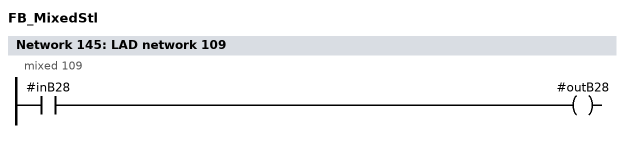
   RUNG wire#powerrail
      Contact( #inB28 )
      Coil( #outB28 )
   END_RUNG
   // the same network as SCL:
   #outB28 := #inB28;
END_REGION

REGION Network 146 (FBD): FBD network 110
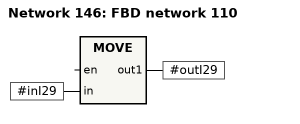
   #outI29 := #inI29;
END_REGION

REGION Network 147 (SCL): SCL network 111
   #tI10 := #inI30 + #cI20;
           IF #inB30 THEN
               #outR10 := #inR10 * 2.0;
           END_IF;
END_REGION

NETWORK
TITLE = STL network 37
      A     #inB36;
      AN    #stB36;
      =     #outB36;

REGION Network 149: LAD network 112
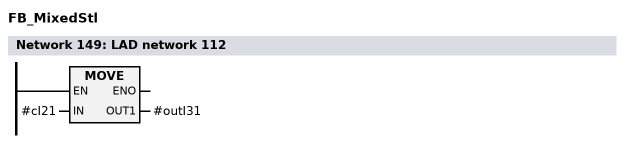
   RUNG wire#powerrail
      Move(in := #cI21, out1 => #outI31)
   END_RUNG
   // the same network as SCL:
   #outI31 := #cI21;
END_REGION

REGION Network 150 (FBD): FBD network 113
   // mixed 113
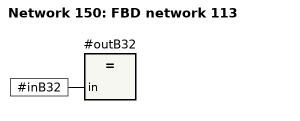
   #outB32 := #inB32;
END_REGION

REGION Network 151 (SCL): SCL network 114
   #tI13 := #inI33 + #cI23;
           IF #inB33 THEN
               #outR13 := #inR13 * 2.0;
           END_IF;
END_REGION

NETWORK
TITLE = STL network 38
      L     #inI37;
      L     #stI37;
      +I;
      T     #outI37;

REGION Network 153: LAD network 115
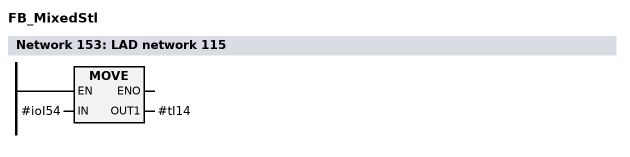
   RUNG wire#powerrail
      Move(in := #ioI54, out1 => #tI14)
   END_RUNG
   // the same network as SCL:
   #tI14 := #ioI54;
END_REGION

REGION Network 154 (FBD): FBD network 116
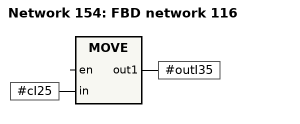
   #outI35 := #cI25;
END_REGION

REGION Network 155 (SCL): SCL network 117
   // mixed 117
   #tI16 := #inI36 + #cI26;
           IF #inB36 THEN
               #outR16 := #inR16 * 2.0;
           END_IF;
END_REGION

NETWORK
TITLE = STL network 39
      L     #inR18;
      L     #tR38;
      *R;
      T     #outR18;  // product

REGION Network 157: LAD network 118
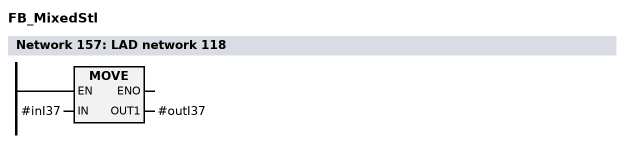
   RUNG wire#powerrail
      Move(in := #inI37, out1 => #outI37)
   END_RUNG
   // the same network as SCL:
   #outI37 := #inI37;
END_REGION

REGION Network 158 (FBD): FBD network 119
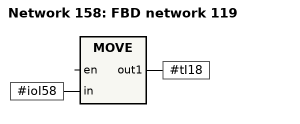
   #tI18 := #ioI58;
END_REGION

REGION Network 159 (SCL): SCL network 120
   #tI19 := #inI39 + #cI29;
           IF #inB39 THEN
               #outR19 := #inR19 * 2.0;
           END_IF;
END_REGION

NETWORK
TITLE = STL network 40
      A     #inB39;
      AN    #stB39;
      =     #outB39;
END_FUNCTION_BLOCK
